(* Munsch response *)
TYPE ET_MUNSCH_RES :
(
	ET_MUNSCH_RES_NOCMD := 0,
	ET_MUNSCH_RES_STARTHEAT := 1,
	ET_MUNSCH_RES_STOPHEAT := 2,
	ET_MUNSCH_RES_ACKHEATSTATUSON := 3,
	ET_MUNSCH_RES_ACKHEATSTATUSOFF := 4,
	ET_MUNSCH_RES_STARTEXTRUDER := 5,
	ET_MUNSCH_RES_STOPEXTRUDER := 6,
	ET_MUNSCH_RES_ACKEXTRUDERSTATUSON := 7,
	ET_MUNSCH_RES_ACKEXTRUDERSTATUSOFF := 8,
	ET_MUNSCH_RES_SETMATERIALTEMP := 9,
	ET_MUNSCH_RES_REQMATERIALREFTEMP := 10,
	ET_MUNSCH_RES_REQMATERIALACTTEMP := 11,
	ET_MUNSCH_RES_SETAIRTEMP := 13,
	ET_MUNSCH_RES_REQAIRREFTEMP := 14,
	ET_MUNSCH_RES_REQAIRACTTEMP := 15,
	ET_MUNSCH_RES_REQSTATUSHEATING := 17,
	ET_MUNSCH_RES_REQSTATUSHEATED := 18,
	ET_MUNSCH_RES_REQSTATUSERROR := 19,
	ET_MUNSCH_RES_CMDERROR := 21

);
END_TYPE

(* stored: Version 1.1.0.1, ProductVersion 3.1.4024.15
   DUT ET_MUNSCH_RES: Id {b8c5236d-1fb3-4432-9715-7792fb826685} *)
